    rq_activate_all_grippers(True)
    # end: URCap Program Node
  end
  $ 56 "zero_ftsensor()"
  zero_ftsensor()
  $ 57 "EXTT"
  $ 58 "Set GRP_3F_Enable=Off"
  set_standard_digital_out(4, False)
  $ 59 "Set BarcodeTrigger=Off"
  set_standard_digital_out(6, False)
  $ 60 "Set GRP_3F_Decap=Off"
  set_standard_digital_out(3, False)
  $ 61 "Set GRP_3F_Cap=Off"
  set_standard_digital_out(2, False)
  $ 62 "Set GRP_3F_Open=Off"
  set_standard_digital_out(5, False)
  $ 63 "PSE_T≔get_tool_free_pose(dir=[0,0,0.150], move_in_base_frame=True)"
  global PSE_T=get_tool_free_pose(dir=[0,0,0.150], move_in_base_frame=True)
  $ 64 "If is_reachable(Base_const, [PSE_T])"
  if (is_reachable(p[0.0,0.0,0.0,0.0,0.0,0.0], [PSE_T])):
    $ 65 "MoveL"
    $ 66 "PSE_T" "breakAfter"
    movel(PSE_T, a=1.2, v=0.15)
  end
  while (True):
    $ 67 "Robot Program"
    $ 68 "MAIN"
    $ 69 "command_manager(external_control='uGO', cond_suspend=(ITM_Manipulated and AMR_AtTarget and AMR_Charging and AMR_Battery<40), cond_unsuspend=(AMR_Battery≟60))"
    command_manager(external_control="uGO", cond_suspend=(ITM_Manipulated  and  AMR_AtTarget  and  AMR_Charging  and  AMR_Battery<40), cond_unsuspend=(AMR_Battery == 60))
    $ 70 "log_state(STATE_Info)"
    log_state(STATE_Info)
    $ 71 "Switch STATE"
    switch_1 = STATE
    $ 72 "Case 1"
    if (1 == switch_1):
      $ 73 "Stopping"
      $ 74 "STATE_Info≔'Stopping'"
      global STATE_Info="Stopping"
      $ 75 "end_freedrive_mode()"
      end_freedrive_mode()
      $ 76 "Set"
      set_tcp(p[0.0,0.0,0.161,3.1415,0.0,0.0])
      $ 77 "PSE_T≔get_tool_free_pose(dir=[0,0,0.150], move_in_base_frame=True)"
      global PSE_T=get_tool_free_pose(dir=[0,0,0.150], move_in_base_frame=True)
      $ 78 "If is_reachable(Base_const, [PSE_T])"
      if (is_reachable(p[0.0,0.0,0.0,0.0,0.0,0.0], [PSE_T])):
        $ 79 "MoveL"
        $ 80 "PSE_T" "breakAfter"
        movel(PSE_T, a=1.2, v=0.15)
      end
      $ 81 "do_transition(keep_rxry=OBJ_Picked, r=0)"
      do_transition(keep_rxry=OBJ_Picked, r=0)
      $ 82 "Decapper"
      $ 83 "Set GRP_3F_Enable=Off"
      set_standard_digital_out(4, False)
      $ 84 "Set BarcodeTrigger=Off"
      set_standard_digital_out(6, False)
      $ 85 "Set GRP_3F_Decap=Off"
      set_standard_digital_out(3, False)
      $ 86 "Set GRP_3F_Cap=Off"
      set_standard_digital_out(2, False)
      $ 87 "Set GRP_3F_Open=Off"
      set_standard_digital_out(5, False)
      $ 90 "Call Sub_AMR_MiR_V3"
      Sub_AMR_MiR_V3()
      $ 91 "If stopping() and AMR_Done"
      if (stopping()  and  AMR_Done):
        $ 92 "STATE≔2"
        global STATE=2
        $ 93 "ugo_update_outputs()"
        ugo_update_outputs()
      end
    elif (2 == switch_1):
      $ 94 "Case 2"
      $ 95 "Stopped"
      $ 96 "STATE_Info≔'Stopped'"
      global STATE_Info="Stopped"
      $ 97 "Call Sub_AMR_MiR_V3"
      Sub_AMR_MiR_V3()
      $ 98 "If CMD_Reset"
      if (CMD_Reset):
        $ 99 "STATE≔3"
        global STATE=3
        $ 100 "ugo_update_outputs()"
        ugo_update_outputs()
      end
    elif (3 == switch_1):
      $ 101 "Case 3"
      $ 102 " Resetting"
      $ 103 "STATE_Info≔'Resetting'"
      global STATE_Info="Resetting"
      $ 104 "uML"
      $ 105 "reset_error()"
      reset_error()
      $ 106 "reset_warning()"
      reset_warning()
      $ 107 "PROCESS_Step≔0"
      global PROCESS_Step=0
      $ 108 "PROCESS_Info≔''"
      global PROCESS_Info=""
      $ 109 "ARM_Referenced≔ False "
      global ARM_Referenced=  False
      $ 110 "WRK_Done≔ False "
      global WRK_Done=  False
      $ 111 "ITM_Prepared≔ False "
      global ITM_Prepared=  False
      $ 112 "ITM_Manipulated≔ False "
      global ITM_Manipulated=  False
      $ 113 "STP≔0"
      global STP=0
      $ 114 "Action≔0"
      global Action=0
      $ 115 "Action_Info≔''"
      global Action_Info=""
      $ 116 "ITM_ID≔0"
      global ITM_ID=0
      $ 117 "JIG≔0"
      global JIG=0
      $ 118 "JIG_Slot≔0"
      global JIG_Slot=0
      $ 119 "Task_info≔''"
      global Task_info=""
      $ 120 "Set"
      set_tcp(p[0.0,0.0,0.161,3.1415,0.0,0.0])
      $ 121 "App"
      $ 122 "'ADD APPLICATION SPECIFIC COMMANDS'"
      # 'ADD APPLICATION SPECIFIC COMMANDS'
      $ 123 "OBJ_Type≔0"
      global OBJ_Type=0
      $ 124 "OBJ_Nbr≔0"
      global OBJ_Nbr=0
      $ 125 "If CNT_Rack_Output≥50"
      if (CNT_Rack_Output >= 50):
        $ 126 "CNT_Rack_Output≔0"
        global CNT_Rack_Output=0
      end
      $ 127 "TASK≔struct(ID=0, NAVI=struct(target=0, footprint=0, protectiveOff=0, dock=0), WORK=struct(ITM_ID_Src=0, JIG_ID_Src=0, OBJ_Nbr_Src=0, ACT_Src=0, ITM_ID_Tgt=0, JIG_ID_Tgt=0, OBJ_Nbr_Tgt=0, ACT_Tgt=0, OBJ_Type=0))"
      global TASK=struct(ID=0, NAVI=struct(target=0, footprint=0, protectiveOff=0, dock=0), WORK=struct(ITM_ID_Src=0, JIG_ID_Src=0, OBJ_Nbr_Src=0, ACT_Src=0, ITM_ID_Tgt=0, JIG_ID_Tgt=0, OBJ_Nbr_Tgt=0, ACT_Tgt=0, OBJ_Type=0))
      $ 128 "Call Sub_AMR_MiR_V3"
      Sub_AMR_MiR_V3()
      $ 129 "If resetting() and AMR_Done"
      if (resetting()  and  AMR_Done):
        $ 130 "STATE≔4"
        global STATE=4
        $ 131 "ugo_update_outputs()"
        ugo_update_outputs()
      end
    elif (4 == switch_1):
      $ 132 "Case 4"
      $ 133 "Idle"
      $ 134 "STATE_Info≔'Idle'"
      global STATE_Info="Idle"
      $ 135 "If CMD_Start"
      if (CMD_Start):
        $ 136 "STATE≔5"
        global STATE=5
        $ 137 "ugo_update_outputs()"
        ugo_update_outputs()
      end
    elif (5 == switch_1):
      $ 138 "Case 5"
      $ 139 "Starting"
      $ 140 "STATE_Info≔'Starting'"
      global STATE_Info="Starting"
      $ 141 "'ADD COMMANDS WHAT TO START WITH'"
      # 'ADD COMMANDS WHAT TO START WITH'
      $ 142 "Call Sub_AMR_MiR_V3"
      Sub_AMR_MiR_V3()
      $ 143 "get ugo data"
      $ 144 "Assign Tasks"
      $ 145 "TASK.ID = ugo_get_task()"
      TASK.ID = ugo_get_task()
      $ 146 "If TASK.ID≟1"
      if (TASK.ID == 1):
        $ 147 "Task_info≔'Charge'"
        global Task_info="Charge"
        $ 148 "Parameters"
        $ 149 "AMR_PosTarget≔1"
        global AMR_PosTarget=1
      else:
        $ 150 "ElseIf TASK.ID≟9"
        if (TASK.ID == 9):
          $ 151 "'Pick Sarstedt Rack from Variable source'"
          # 'Pick Sarstedt Rack from Variable source'
          $ 152 "Task_info≔'Navigate to Target'"
          global Task_info="Navigate to Target"
          $ 153 "Parameters"
          $ 154 "AMR_PosTarget≔UGO.read_input('00','ITM_ID')"
          global AMR_PosTarget=UGO.read_input("00","ITM_ID")
        else:
          $ 155 "ElseIf TASK.ID≟10"
          if (TASK.ID == 10):
            $ 156 "'Pick Sarstedt Rack from Variable source'"
            # 'Pick Sarstedt Rack from Variable source'
            $ 157 "Task_info≔'Pick Rack'"
            global Task_info="Pick Rack"
            $ 158 "AMR_PosTarget≔2"
            global AMR_PosTarget=2
            $ 159 "Parameters"
            $ 160 "ITM_ID≔UGO.read_input('00','ITM_ID')"
            global ITM_ID=UGO.read_input("00","ITM_ID")
            $ 161 "JIG≔UGO.read_input('00','JIG_ID')"
            global JIG=UGO.read_input("00","JIG_ID")
            $ 162 "OBJ_Type≔3"
            global OBJ_Type=3
          else:
            $ 164 "ElseIf TASK.ID≟11"
            if (TASK.ID == 11):
              $ 165 "'Place Sarstedt Rack on Variable target'"
              # 'Place Sarstedt Rack on Variable target'
              $ 166 "Task_info≔'Place Rack'"
              global Task_info="Place Rack"
              $ 167 "AMR_PosTarget≔2"
              global AMR_PosTarget=2
              $ 168 "Parameters"
              $ 169 "ITM_ID≔UGO.read_input('00','ITM_ID')"
              global ITM_ID=UGO.read_input("00","ITM_ID")
              $ 170 "JIG≔UGO.read_input('00','JIG_ID')"
              global JIG=UGO.read_input("00","JIG_ID")
              $ 171 "OBJ_Type≔3"
              global OBJ_Type=3
            else:
              $ 173 "ElseIf TASK.ID≟12"
              if (TASK.ID == 12):
                $ 174 "Task_info≔'Decapping'"
                global Task_info="Decapping"
                $ 175 "Parameters"
                $ 176 "ITM_ID≔1"
                global ITM_ID=1
                $ 177 "OBJ_Type≔2"
                global OBJ_Type=2
                $ 178 "JIG≔2"
                global JIG=2
                $ 179 "AMR_PosTarget≔AMR_PosActual"
                global AMR_PosTarget=AMR_PosActual
                $ 180 "PRC_TubCounter≔0"
                global PRC_TubCounter=0
              else:
                $ 181 "ElseIf TASK.ID≟13"
                if (TASK.ID == 13):
                  $ 182 "Task_info≔'Empty racks'"
                  global Task_info="Empty racks"
                  $ 183 "Parameters"
                  $ 184 "ITM_ID≔1"
                  global ITM_ID=1
                  $ 185 "AMR_PosTarget≔AMR_PosActual"
                  global AMR_PosTarget=AMR_PosActual
                else:
                  $ 186 "ElseIf TASK.ID≟14"
                  if (TASK.ID == 14):
                    $ 187 "Task_info≔'Decap'"
                    global Task_info="Decap"
                    $ 188 "Parameters"
                    $ 189 "ITM_ID≔1"
                    global ITM_ID=1
                    $ 190 "OBJ_Type≔2"
                    global OBJ_Type=2
                    $ 191 "JIG≔7"
                    global JIG=7
                    $ 192 "AMR_PosTarget≔AMR_PosActual"
                    global AMR_PosTarget=AMR_PosActual
                  else:
                    $ 193 "ElseIf TASK.ID≟99"
                    if (TASK.ID == 99):
                      $ 194 "Task_info≔'Decapping and barcode alignment'"
                      global Task_info="Decapping and barcode alignment"
                      $ 195 "Parameters"
                      $ 196 "PRC_TubNumber≔UGO.read_input('00','TubesNb')"
                      global PRC_TubNumber=UGO.read_input("00","TubesNb")
                      $ 197 "PRC_TubCounter≔0"
                      global PRC_TubCounter=0
                      $ 198 "ITM_ID≔1"
                      global ITM_ID=1
                      $ 199 "AMR_PosTarget≔AMR_PosActual"
                      global AMR_PosTarget=AMR_PosActual
                    else:
                      $ 208 "ElseIf TASK.ID≟15"
                      if (TASK.ID == 15):
                        $ 209 "Task_info≔'Unoad Centrifuge'"
                        global Task_info="Unoad Centrifuge"
                        $ 210 "Parameters"
                        $ 211 "PRC_RackCounter≔0"
                        global PRC_RackCounter=0
                        $ 212 "TASK.WORK.ITM_ID_Src=2"
                        TASK.WORK.ITM_ID_Src=2
                        $ 213 "TASK.WORK.ITM_ID_Tgt=1"
                        TASK.WORK.ITM_ID_Tgt=1
                        $ 214 "AMR_PosTarget≔4"
                        global AMR_PosTarget=4
                        $ 215 "AMR_FootprintID≔1"
                        global AMR_FootprintID=1
                      else:
                        $ 234 "Else" "noBreak"
                        $ 235 "set_error(ERROR_WRONG_ORDER)"
                        set_error(ERROR_WRONG_ORDER)
                      end
                    end
                  end
                end
              end
            end
          end
        end
      end
      $ 236 "test ugo"
      $ 237 "Wait: 0.2"
      sleep(0.2)
      $ 238 "ugo_update_outputs()"
      ugo_update_outputs()
      $ 239 "If starting() and AMR_Done"
      if (starting()  and  AMR_Done):
        $ 240 "log_message(Task_info, 'New Task: ')"
        log_message(Task_info, "New Task: ")
        $ 241 "log_message(to_str(TASK.ID), 'Task_ID: ')"
        log_message(to_str(TASK.ID), "Task_ID: ")
        $ 242 "do_transition(keep_rxry=OBJ_Picked)"
        do_transition(keep_rxry=OBJ_Picked)
        $ 243 "STATE≔6"
        global STATE=6
        $ 244 "ugo_update_outputs()"
        ugo_update_outputs()
      end
    elif (6 == switch_1):
      $ 245 "Case 6"
      $ 246 "Execute"
      $ 247 "STATE_Info≔'Execute'"
      global STATE_Info="Execute"
      $ 248 "If  not CMD_Hold and not CMD_Suspend"
      global thread_flag_248=0
      thread Thread_if_248():
        $ 249 "Switch PROCESS_Step"
        switch_2 = PROCESS_Step
        $ 250 "Case 0"
        if (0 == switch_2):
          $ 251 "PROCESS_Info≔'process control'"
          global PROCESS_Info="process control"
          $ 252 "log_process(PROCESS_Info)"
          log_process(PROCESS_Info)
          $ 253 "process control"
          $ 254 "If  not AMR_AtTarget"
          if (  not  AMR_AtTarget):
            $ 255 "PROCESS_Step≔1"
            global PROCESS_Step=1
          else:
            $ 256 "ElseIf (( not ITM_Prepared and  not WRK_Done) or (ITM_Prepared and WRK_Done))"
            if (((  not  ITM_Prepared  and    not  WRK_Done)  or  (ITM_Prepared  and  WRK_Done))):
              $ 257 "PROCESS_Step≔2"
              global PROCESS_Step=2
            else:
              $ 258 "ElseIf  not WRK_Done"
              if (  not  WRK_Done):
                $ 259 "PROCESS_Step≔3"
                global PROCESS_Step=3
              else:
                $ 260 "Else" "noBreak"
                $ 261 "task finished"
                $ 262 "PROCESS_Info≔''"
                global PROCESS_Info=""
                $ 263 "STATE≔7"
                global STATE=7
                $ 264 "ugo_update_outputs()"
                ugo_update_outputs()
              end
            end
          end
        elif (1 == switch_2):
          $ 265 "Case 1"
          $ 266 "navigate"
          $ 267 "'MOVING THE uML'"
          # 'MOVING THE uML'
          $ 268 "PROCESS_Info≔'move to target'"
          global PROCESS_Info="move to target"
          $ 269 "log_process(PROCESS_Info)"
          log_process(PROCESS_Info)
          $ 270 "If TASK.ID≟1"
          if (TASK.ID == 1):
            $ 271 "Action≔51"
            global Action=51
          else:
            $ 272 "Else" "noBreak"
            $ 273 "Action≔52"
            global Action=52
          end
          $ 274 "Call Sub_AMR_MiR_V3"
          Sub_AMR_MiR_V3()
          $ 275 "If AMR_Done"
          if (AMR_Done):
            $ 276 "PROCESS_Step≔0"
            global PROCESS_Step=0
          end
        elif (2 == switch_2):
          $ 277 "Case 2"
          $ 278 "prepare"
          $ 279 "'THINGS THAT HAVE TO BE DONE ONCE IN A SEQUENCE,WORKFLOW'"
          # 'THINGS THAT HAVE TO BE DONE ONCE IN A SEQUENCE,WORKFLOW'
          $ 280 "PROCESS_Info≔'prepare for work'"
          global PROCESS_Info="prepare for work"
          $ 281 "log_process(PROCESS_Info)"
          log_process(PROCESS_Info)
          $ 282 "If TASK.WORK.ITM_ID_Src>1"
          if (TASK.WORK.ITM_ID_Src>1):
            $ 283 "ITM_ID≔TASK.WORK.ITM_ID_Src"
            global ITM_ID=TASK.WORK.ITM_ID_Src
          else:
            $ 284 "ElseIf TASK.WORK.ITM_ID_Tgt>1"
            if (TASK.WORK.ITM_ID_Tgt>1):
              $ 285 "ITM_ID≔TASK.WORK.ITM_ID_Tgt"
              global ITM_ID=TASK.WORK.ITM_ID_Tgt
            end
          end
          $ 286 "If  not ARM_Referenced and (ITM_ID≠0)"
          if (  not  ARM_Referenced  and  (ITM_ID != 0)):
            $ 287 "STP≔1"
            global STP=1
          else:
            $ 288 "ElseIf ARM_Referenced or (ITM_ID≟0)"
            if (ARM_Referenced  or  (ITM_ID == 0)):
              $ 289 "STP≔2"
              global STP=2
            end
          end
          $ 290 "Switch STP"
          switch_3 = STP
          $ 291 "Case 1"
          if (1 == switch_3):
            $ 292 "reference"
            $ 293 "STP_Info≔'reference at target position'"
            global STP_Info="reference at target position"
            $ 294 "log_step(STP_Info)"
            log_step(STP_Info)
            $ 295 "If ITM_ID≟1"
            if (ITM_ID == 1):
              $ 296 "CAM_Done≔ True "
              global CAM_Done=  True
            else:
              $ 297 "Else" "noBreak"
              $ 298 "Action≔131"
              global Action=131
              $ 299 "Call Sub_Vision_V18"
              Sub_Vision_V18()
            end
            $ 301 "If CAM_Done and  not ERROR.FLAG"
            if (CAM_Done  and    not  ERROR.FLAG):
              $ 302 "log_step('ARM referenced')"
              log_step("ARM referenced")
              $ 303 "ARM_Referenced≔ True "
              global ARM_Referenced=  True
            end
          elif (2 == switch_3):
            $ 304 "Case 2"
            $ 305 "manipulate"
            $ 306 "STP_Info≔'manipulate item'"
            global STP_Info="manipulate item"
            $ 307 "log_step(STP_Info)"
            log_step(STP_Info)
            $ 308 "'In case pressing button is needed'"
            # 'In case pressing button is needed'
            $ 309 "If found_in_list(ITM_ID, ITM_ID_List)"
            if (found_in_list(ITM_ID, ITM_ID_List)):
              $ 310 "Switch ITM_ID"
              switch_4 = ITM_ID
              $ 311 "Case 0"
              if (0 == switch_4):
                $ 312 "ITM_Manipulated≔ not ITM_Manipulated"
                global ITM_Manipulated=  not  ITM_Manipulated
              elif (1 == switch_4):
                $ 313 "Case 1"
                $ 314 "ITM_Manipulated≔ not ITM_Manipulated"
                global ITM_Manipulated=  not  ITM_Manipulated
              elif (2 == switch_4):
                $ 315 "Case 2"
              else:
                $ 325 "Default Case"
                $ 326 "ITM_Manipulated≔ not ITM_Manipulated"
                global ITM_Manipulated=  not  ITM_Manipulated
              end
            end
          end
          $ 327 "ITM_Prepared≔(ITM_Manipulated or  not found_in_list(ITM_ID, ITM_ID_List)) and (ARM_Referenced or ITM_ID≟0) and  not WRK_Done"
          global ITM_Prepared=(ITM_Manipulated  or    not  found_in_list(ITM_ID, ITM_ID_List))  and  (ARM_Referenced  or  ITM_ID == 0)  and    not  WRK_Done
          $ 328 "STP≔0"
          global STP=0
          $ 329 "STP_Info≔''"
          global STP_Info=""
          $ 330 "PROCESS_Step≔0"
          global PROCESS_Step=0
        elif (3 == switch_2):
          $ 331 "Case 3"
          $ 332 "work"
          $ 333 "'ADD EVERY MACHINE, OBJECT, STATION TO WORK ON'"
          # 'ADD EVERY MACHINE, OBJECT, STATION TO WORK ON'
          $ 334 "Switch ITM_ID"
          switch_3 = ITM_ID
          $ 335 "Case 1"
          if (1 == switch_3):
            $ 336 "uLM"
            $ 337 "If TASK.ID≟12"
            if (TASK.ID == 12):
            else:
              $ 365 "ElseIf TASK.ID≟10"
              if (TASK.ID == 10):
                $ 366 "Pick Rack"
                $ 367 "Action≔131"
                global Action=131
                $ 368 "Call Sub_Vision_V18"
                Sub_Vision_V18()
                $ 369 "Action≔1"
                global Action=1
                $ 370 "Call Sub_Action_V4"
                Sub_Action_V4()
                $ 371 "PROCESS_Step≔0"
                global PROCESS_Step=0
                $ 372 "WRK_Done≔ True "
                global WRK_Done=  True
              else:
                $ 373 "ElseIf TASK.ID≟11"
                if (TASK.ID == 11):
                  $ 374 "Place Rack"
                  $ 375 "Action≔2"
                  global Action=2
                  $ 376 "Call Sub_Action_V4"
                  Sub_Action_V4()
                  $ 377 "PROCESS_Step≔0"
                  global PROCESS_Step=0
                  $ 378 "WRK_Done≔ True "
                  global WRK_Done=  True
                else:
                  $ 379 "ElseIf TASK.ID≟13"
                  if (TASK.ID == 13):
                    $ 380 "empty racks"
                    $ 381 "pick"
                    $ 382 "Action≔1"
                    global Action=1
                    $ 383 "JIG≔4"
                    global JIG=4
                    $ 384 "If PRC_TubCounter%4≟0"
                    if (PRC_TubCounter%4 == 0):
                      $ 385 "JIG_Slot≔4"
                      global JIG_Slot=4
                    else:
                      $ 386 "Else" "noBreak"
                      $ 387 "JIG_Slot≔PRC_TubCounter%4"
                      global JIG_Slot=PRC_TubCounter%4
                    end
                    $ 388 "OBJ_Nbr≔ceil(PRC_TubCounter/4)"
                    global OBJ_Nbr=ceil(PRC_TubCounter/4)
                    $ 389 "OBJ_Type≔2"
                    global OBJ_Type=2
                    $ 390 "Call Sub_Action_V4"
                    Sub_Action_V4()
                    $ 391 "If OBJ_Picked"
                    if (OBJ_Picked):
                      $ 392 "Action≔2"
                      global Action=2
                      $ 393 "JIG≔3"
                      global JIG=3
                      $ 394 "JIG_Slot≔1"
                      global JIG_Slot=1
                      $ 395 "CNT_Rack_Output≔CNT_Rack_Output + 1"
                      global CNT_Rack_Output=CNT_Rack_Output + 1
                      $ 396 "OBJ_Nbr≔CNT_Rack_Output"
                      global OBJ_Nbr=CNT_Rack_Output
                      $ 397 "Call Sub_Action_V4"
                      Sub_Action_V4()
                      $ 398 "If  not ERROR.FLAG"
                      if (  not  ERROR.FLAG):
                        $ 399 "PRC_TubCounter≔PRC_TubCounter - 1"
                        global PRC_TubCounter=PRC_TubCounter - 1
                      end
                    end
                    $ 400 "If CNT_Rack_Output≥50 or PRC_TubCounter≤0"
                    if (CNT_Rack_Output >= 50  or  PRC_TubCounter <= 0):
                      $ 401 "PROCESS_Step≔0"
                      global PROCESS_Step=0
                      $ 402 "WRK_Done≔ True "
                      global WRK_Done=  True
                    end
                  else:
                    $ 403 "ElseIf TASK.ID≟14"
                    if (TASK.ID == 14):
                      $ 407 "JIG≔7"
                      global JIG=7
                      $ 408 "Action≔151"
                      global Action=151
                      $ 409 "Call Sub_Vision_V18"
                      Sub_Vision_V18()
                      $ 410 "PRC_CntDetect≔0"
                      global PRC_CntDetect=0
                      $ 412 "If CAM_Result.length()>0"
                      if (CAM_Result.length()>0):
                        $ 413 "samples≔ True "
                        global samples=  True
                      else:
                        $ 414 "Else" "noBreak"
                        $ 415 "samples≔ False "
                        global samples=  False
                      end
                      $ 416 "Loop samples≟ True "
                      while (samples ==   True  ):
                        $ 417 "Action≔1"
                        global Action=1
                        $ 418 "ITM_ID≔1"
                        global ITM_ID=1
                        $ 419 "JIG≔2"
                        global JIG=2
                        $ 420 "OBJ_Type≔2"
                        global OBJ_Type=2
                        $ 421 "JIG_Slot≔CAM_Result[PRC_CntDetect]"
                        global JIG_Slot=CAM_Result[PRC_CntDetect]
                        $ 422 "OBJ_Nbr≔CAM_Result[PRC_CntDetect]"
                        global OBJ_Nbr=CAM_Result[PRC_CntDetect]
                        $ 423 "Call Sub_Action_V4"
                        Sub_Action_V4()
                        $ 437 "JIG≔2"
                        global JIG=2
                        $ 438 "Action≔2"
                        global Action=2
                        $ 439 "OBJ_Nbr≔CAM_Result[PRC_CntDetect]"
                        global OBJ_Nbr=CAM_Result[PRC_CntDetect]
                        $ 440 "JIG_Slot≔CAM_Result[PRC_CntDetect]"
                        global JIG_Slot=CAM_Result[PRC_CntDetect]
                        $ 441 "OBJ_Type≔2"
                        global OBJ_Type=2
                        $ 442 "Call Sub_Action_V4"
                        Sub_Action_V4()
                        $ 443 "PRC_CntDetect≔PRC_CntDetect+1"
                        global PRC_CntDetect=PRC_CntDetect+1
                        $ 444 "If CAM_Result.length()<=PRC_CntDetect"
                        if (CAM_Result.length()<=PRC_CntDetect):
                          $ 445 "samples≔ False "
                          global samples=  False
                        end
                      end
                    end
                  end
                end
              end
            end
          elif (2 == switch_3):
            $ 446 "Case 2"
          elif (20 == switch_3):
            $ 488 "Case 20"
          else:
            $ 550 "Default Case"
            $ 551 "WRK_Done≔ True "
            global WRK_Done=  True
            $ 552 "PROCESS_Step≔0"
            global PROCESS_Step=0
          end
        end
        thread_flag_248 = 1
      end
      if (  not  CMD_Hold and not CMD_Suspend):
        global thread_handler_248=run Thread_if_248()
        while (thread_flag_248 == 0):
          if not(  not  CMD_Hold and not CMD_Suspend):
            kill thread_handler_248
            thread_flag_248 = 2
          else:
            sync()
          end
        end
      else:
        thread_flag_248 = 2
      end
      $ 553 "If CMD_Hold"
      if (CMD_Hold):
        $ 554 "STATE≔9"
        global STATE=9
        $ 555 "ugo_update_outputs()"
        ugo_update_outputs()
      else:
        $ 556 "ElseIf CMD_Suspend"
        if (CMD_Suspend):
          $ 557 "STATE≔12"
          global STATE=12
          $ 558 "ugo_update_outputs()"
          ugo_update_outputs()
        end
      end
    elif (7 == switch_1):
      $ 559 "Case 7"
      $ 560 "Completing"
      $ 561 "STATE_Info≔'Completing'"
      global STATE_Info="Completing"
      $ 562 "'ADD COMMANDS FOR COMPLETING THE PROCESS'"
      # 'ADD COMMANDS FOR COMPLETING THE PROCESS'
      $ 563 "do_transition(keep_rxry=OBJ_Picked)"
      do_transition(keep_rxry=OBJ_Picked)
      $ 564 "Call Sub_AMR_MiR_V3"
      Sub_AMR_MiR_V3()
      $ 565 "If completing() and AMR_Done"
      if (completing()  and  AMR_Done):
        $ 566 "STATE≔8"
        global STATE=8
        $ 567 "ugo_update_outputs()"
        ugo_update_outputs()
      end
    elif (8 == switch_1):
      $ 568 "Case 8"
      $ 569 "Complete"
      $ 570 "STATE_Info≔'Complete'"
      global STATE_Info="Complete"
      $ 571 "If CMD_Reset"
      if (CMD_Reset):
        $ 572 "STATE≔3"
        global STATE=3
        $ 573 "ugo_update_outputs()"
        ugo_update_outputs()
      end
    elif (9 == switch_1):
      $ 574 "Case 9"
      $ 575 "Holding"
      $ 576 "STATE_Info≔'Holding'"
      global STATE_Info="Holding"
      $ 577 "stopl(0.5)"
      stopl(0.5)
      $ 578 "Call Sub_AMR_MiR_V3"
      Sub_AMR_MiR_V3()
      $ 579 "If holding() and AMR_Done"
      if (holding()  and  AMR_Done):
        $ 580 "STATE≔10"
        global STATE=10
        $ 581 "ugo_update_outputs()"
        ugo_update_outputs()
      end
    elif (10 == switch_1):
      $ 582 "Case 10"
      $ 583 "Held"
      $ 584 "STATE_Info≔'Held'"
      global STATE_Info="Held"
      $ 585 "If CMD_Unhold"
      if (CMD_Unhold):
        $ 586 "end_freedrive_mode()"
        end_freedrive_mode()
        $ 587 "STATE≔11"
        global STATE=11
        $ 588 "ugo_update_outputs()"
        ugo_update_outputs()
      else:
        $ 589 "ElseIf FNC_Freedrive"
        if (FNC_Freedrive):
          $ 590 "freedrive_mode()"
          freedrive_mode()
        else:
          $ 591 "Else" "noBreak"
          $ 592 "end_freedrive_mode()"
          end_freedrive_mode()
        end
      end
    elif (11 == switch_1):
      $ 593 "Case 11"
      $ 594 "Unholding"
      $ 595 "STATE_Info≔'Unholding'"
      global STATE_Info="Unholding"
      $ 596 "Clearing"
      $ 597 "Switch ERROR.ID"
      switch_2 = ERROR.ID
      $ 598 "Case 1002"
      if (1002 == switch_2):
        $ 599 "AMR_AtTarget≔ False "
        global AMR_AtTarget=  False
        $ 600 "ARM_Referenced≔ False "
        global ARM_Referenced=  False
        $ 601 "ITM_Prepared≔ False "
        global ITM_Prepared=  False
        $ 602 "PROCESS_Step≔1"
        global PROCESS_Step=1
      elif (2007 == switch_2):
        $ 603 "Case 2007"
        $ 604 "PROCESS_Step≔1"
        global PROCESS_Step=1
      end
      $ 605 "reset_error()"
      reset_error()
      $ 606 "reset_warning()"
      reset_warning()
      $ 607 "OBJ_Picked≔gripper_has_object()"
      global OBJ_Picked=gripper_has_object()
      $ 608 "Call Sub_AMR_MiR_V3"
      Sub_AMR_MiR_V3()
      $ 609 "If unholding() and AMR_Done"
      if (unholding()  and  AMR_Done):
        $ 610 "STATE≔6"
        global STATE=6
        $ 611 "ugo_update_outputs()"
        ugo_update_outputs()
      end
    elif (12 == switch_1):
      $ 612 "Case 12"
      $ 613 "Suspending"
      $ 614 "STATE_Info≔'Suspending'"
      global STATE_Info="Suspending"
      $ 615 "PROCESS_Info≔str_cat(PROCESS_Info, ' suspended')"
      global PROCESS_Info=str_cat(PROCESS_Info, " suspended")
      $ 616 "If suspending()"
      if (suspending()):
        $ 617 "STATE≔13"
        global STATE=13
        $ 618 "ugo_update_outputs()"
        ugo_update_outputs()
      end
    elif (13 == switch_1):
      $ 619 "Case 13"
      $ 620 "Suspended"
      $ 621 "STATE_Info≔'Suspended'"
      global STATE_Info="Suspended"
      $ 622 "Call Sub_AMR_MiR_V3"
      Sub_AMR_MiR_V3()
      $ 623 "If CMD_Unsuspend"
      if (CMD_Unsuspend):
        $ 624 "STATE≔14"
        global STATE=14
        $ 625 "ugo_update_outputs()"
        ugo_update_outputs()
      end
    elif (14 == switch_1):
      $ 626 "Case 14"
      $ 627 "Unsuspending"
      $ 628 "STATE_Info≔'Unsuspending'"
      global STATE_Info="Unsuspending"
      $ 629 "PROCESS_Step≔0"
      global PROCESS_Step=0
      $ 630 "If unsuspending()"
      if (unsuspending()):
        $ 631 "STATE≔6"
        global STATE=6
        $ 632 "ugo_update_outputs()"
        ugo_update_outputs()
      end
    elif (15 == switch_1):
      $ 633 "Case 15"
      $ 634 "Aborting"
      $ 635 "STATE_Info≔'Aborting'"
      global STATE_Info="Aborting"
      $ 636 "If aborting()"
      if (aborting()):
        $ 637 "STATE≔16"
        global STATE=16
        $ 638 "ugo_update_outputs()"
        ugo_update_outputs()
      end
    elif (16 == switch_1):
      $ 639 "Case 16"
      $ 640 "Aborted"
      $ 641 "STATE_Info≔'Aborted'"
      global STATE_Info="Aborted"
      $ 642 "If CMD_Clear"
      if (CMD_Clear):
        $ 643 "STATE≔17"
        global STATE=17
        $ 644 "ugo_update_outputs()"
        ugo_update_outputs()
      end
    elif (17 == switch_1):
      $ 645 "Case 17"
      $ 646 "Clearing"
      $ 647 "STATE_Info≔'Clearing'"
      global STATE_Info="Clearing"
      $ 648 "Clearing"
      $ 649 "reset_warning()"
      reset_warning()
      $ 650 "reset_error()"
      reset_error()
      $ 651 "If clearing()"
      if (clearing()):
        $ 652 "STATE≔2"
        global STATE=2
        $ 653 "ugo_update_outputs()"
        ugo_update_outputs()
      end
    end
    $ 654 "log_state(STATE_Info)"
    log_state(STATE_Info)
    $ 655 "log_warning(WARNING.MSG)"
    log_warning(WARNING.MSG)
    $ 656 "log_error(ERROR.MSG)"
    log_error(ERROR.MSG)
    $ 657 "Times"
    $ 658 "Switch STATE"
    switch_1 = STATE
    $ 659 "Case 1"
    if (1 == switch_1):
      $ 660 "TM_St_Stopping≔get_time(STATE_Times[STATE-1])"
      global TM_St_Stopping=get_time(STATE_Times[STATE-1])
    elif (2 == switch_1):
      $ 661 "Case 2"
      $ 662 "TM_St_Stopped≔get_time(STATE_Times[STATE-1])"
      global TM_St_Stopped=get_time(STATE_Times[STATE-1])
    elif (3 == switch_1):
      $ 663 "Case 3"
      $ 664 "TM_St_Resetting≔get_time(STATE_Times[STATE-1])"
      global TM_St_Resetting=get_time(STATE_Times[STATE-1])
    elif (4 == switch_1):
      $ 665 "Case 4"
      $ 666 "TM_St_Idle≔get_time(STATE_Times[STATE-1])"
      global TM_St_Idle=get_time(STATE_Times[STATE-1])
    elif (5 == switch_1):
      $ 667 "Case 5"
      $ 668 "TM_St_Starting≔get_time(STATE_Times[STATE-1])"
      global TM_St_Starting=get_time(STATE_Times[STATE-1])
    elif (6 == switch_1):
      $ 669 "Case 6"
      $ 670 "TM_St_Execute≔get_time(STATE_Times[STATE-1])"
      global TM_St_Execute=get_time(STATE_Times[STATE-1])
    elif (7 == switch_1):
      $ 671 "Case 7"
      $ 672 "TM_St_Completin≔get_time(STATE_Times[STATE-1])"
      global TM_St_Completin=get_time(STATE_Times[STATE-1])
    elif (8 == switch_1):
      $ 673 "Case 8"
      $ 674 "TM_St_Complete≔get_time(STATE_Times[STATE-1])"
      global TM_St_Complete=get_time(STATE_Times[STATE-1])
    elif (9 == switch_1):
      $ 675 "Case 9"
      $ 676 "TM_St_Holding≔get_time(STATE_Times[STATE-1])"
      global TM_St_Holding=get_time(STATE_Times[STATE-1])
    elif (10 == switch_1):
      $ 677 "Case 10"
      $ 678 "TM_St_Held≔get_time(STATE_Times[STATE-1])"
      global TM_St_Held=get_time(STATE_Times[STATE-1])
    elif (11 == switch_1):
      $ 679 "Case 11"
      $ 680 "TM_St_Unholding≔get_time(STATE_Times[STATE-1])"
      global TM_St_Unholding=get_time(STATE_Times[STATE-1])
    elif (12 == switch_1):
      $ 681 "Case 12"
      $ 682 "TM_St_Suspendin≔get_time(STATE_Times[STATE-1])"
      global TM_St_Suspendin=get_time(STATE_Times[STATE-1])
    elif (13 == switch_1):
      $ 683 "Case 13"
      $ 684 "TM_St_Suspended≔get_time(STATE_Times[STATE-1])"
      global TM_St_Suspended=get_time(STATE_Times[STATE-1])
    elif (14 == switch_1):
      $ 685 "Case 14"
      $ 686 "TM_St_Unsuspend≔get_time(STATE_Times[STATE-1])"
      global TM_St_Unsuspend=get_time(STATE_Times[STATE-1])
    elif (15 == switch_1):
      $ 687 "Case 15"
      $ 688 "TM_St_Aborting≔get_time(STATE_Times[STATE-1])"
      global TM_St_Aborting=get_time(STATE_Times[STATE-1])
    elif (16 == switch_1):
      $ 689 "Case 16"
      $ 690 "TM_St_Aborted≔get_time(STATE_Times[STATE-1])"
      global TM_St_Aborted=get_time(STATE_Times[STATE-1])
    elif (17 == switch_1):
      $ 691 "Case 17"
      $ 692 "TM_St_Clearing≔get_time(STATE_Times[STATE-1])"
      global TM_St_Clearing=get_time(STATE_Times[STATE-1])
    end
    $ 694 "Wait: 0.1"
    sleep(0.1)
  end
end
